Staubli VAL3: setAnaOutput.pgx

public program setAnaOutput(num x_nIndex, num x_nValue, num& x_nResult)
  local string l_sDesc
  local string l_sPath
//写模拟输出 aOutput[x_nIndex]
//返回码 x_nResult: 0=正常  -1=索引越界  -2=该路未绑定物理通道(aioSet 会 runtime error，已提前拦截)
//注意：aOutput 还没有 link（未做物理 IO 导入），此时写入不会作用到任何物理通道，
//      必须先在 SRS 里完成物理 IO 导入，见 docs/05-IO绑定方法.md
begin
  x_nResult=0

  //越界检查：合法下标 0..size(aOutput)-1（手册 2.5.4，第31页 num size(*)）
  if (x_nIndex<0) or (x_nIndex>=size(aOutput))
    x_nResult=-1
    return
  endIf

  //手册 3.6.1（第63页）：未 link 的 aio 参与运算会 runtime error，所以必须先 ioStatus
  if ioStatus(aOutput[x_nIndex],l_sDesc,l_sPath)<0
    x_nResult=-2
    return
  endIf

  aioSet(aOutput[x_nIndex],x_nValue)
end
